Yaskawa INFORM job: CONFPRO.JBI

/JOB
//NAME CONFPRO
//POS
///NPOS 8,0,0,0,0,0
///TOOL 9
///POSTYPE PULSE
///PULSE
C00000=0,-10240,0,-34475,0,0,22983
C00001=189440,-10240,-218340,-34475,310272,-116053,22983
C00002=-189440,-61440,218340,34475,-425188,116053,114916
C00003=10240,20480,-45966,57458,-68949,-40619,-34475
C00004=-174080,46080,195356,-103424,205699,52224,-51712
C00005=-174080,46080,195356,-103424,205699,52224,-51712
C00006=189440,-10240,-218340,-34475,310272,-116053,22983
C00007=-189440,-61440,218340,34475,-425188,116053,114916
//INST
<volatile>
///COMM Generated using RoboDK
///ATTR SC,RW
///GROUP1 RB1
NOP
'Program generated by RoboDK v
'6.0.7 for Yaskawa Motoman CSD
'A10F on XX/XX/XXXX 18:00:00
'Using nominal kinematics.
'Using Frame S (targets wrt ba
'se):
'1234.6,-98.8,50.5,0.0,0.0,30.
'0
'Tool Tool S should be close t
'o:
'10.0,20.0,150.0,0.0,0.0,0.0
MOVL C00000 V=100.0
MOVL C00001 V=100.0
MOVL C00002 V=100.0
MOVJ C00003 VJ=50.00
MOVJ C00004 VJ=50.00
MOVC C00005 V=100.0
MOVC C00006 V=100.0
MOVC C00007 V=100.0
END
